(* IEC 61131-3 sources: llm-plc-st-eval/data/definitivo/qwen2.5-coder_14b/I5/zero_shot, 3 files *)

(* ---- ejec_1.st ---- *)
```pascal
FUNCTION_BLOCK FB_Clasificadora
VAR_INPUT
    sensorPresencia : BOOL; // Sensor de presencia de pieza
    sensorAltura : BOOL;    // Sensor de altura de pieza
END_VAR

VAR_OUTPUT
    banda : BOOL;          // Salida para activar la banda
    piston : BOOL;         // Salida para activar el pistón
END_VAR

VAR
    nAltas : INT := 0;      // Contador de piezas altas
    nBajas : INT := 0;      // Contador de piezas bajas
    timer1 : TON;           // Timer para el tiempo de espera (2s)
    timer2 : TON;           // Timer para el tiempo de activación del pistón (1s)
    estado : INT := 0;      // Estado de la máquina de estados
END_VAR

// Máquina de estados
CASE estado OF
    0: // Estado inicial
        banda := TRUE; // La banda funciona continuamente
        IF sensorPresencia THEN
            estado := 1; // Detectada pieza, iniciar temporizador
            timer1(IN := TRUE, PT := T#2S); // Iniciar temporizador de 2s
        END_IF

    1: // Esperando que la pieza llegue al desviador
        IF timer1.Q THEN
            IF sensorAltura THEN
                estado := 2; // Pieza alta, activar pistón
                timer2(IN := TRUE, PT := T#1S); // Iniciar temporizador de 1s
                nAltas := nAltas + 1; // Incrementar contador de piezas altas
            ELSE
                estado := 0; // Pieza baja, continuar
                nBajas := nBajas + 1; // Incrementar contador de piezas bajas
            END_IF
        END_IF

    2: // Activando el pistón
        piston := TRUE;
        IF timer2.Q THEN
            piston := FALSE; // Desactivar pistón
            estado := 0; // Volver al estado inicial
        END_IF

    ELSE
        estado := 0; // Estado desconocido, volver al inicial
END_CASE
```

(* ---- ejec_2.st ---- *)
```iec
FUNCTION_BLOCK FB_Clasificadora
VAR_INPUT
    sensorPresencia : BOOL; // Sensor de presencia de pieza
    sensorAltura : BOOL;    // Sensor de altura de pieza
END_VAR

VAR_OUTPUT
    banda : BOOL;          // Salida para activar la banda
    piston : BOOL;         // Salida para activar el pistón
    nAltas : INT;          // Contador de piezas altas
    nBajas : INT;          // Contador de piezas bajas
END_VAR

VAR
    timer1 : TON;           // Timer para esperar 2 segundos
    timer2 : TON;           // Timer para activar el pistón durante 1 segundo
    piezaDetectada : BOOL;  // Bandera para detectar pieza
END_VAR

// Inicialización de variables
IF NOT piezaDetectada THEN
    timer1(IN := FALSE);
    timer2(IN := FALSE);
    piston := FALSE;
END_IF

// Detectar pieza
IF sensorPresencia AND NOT piezaDetectada THEN
    piezaDetectada := TRUE;
    timer1(IN := TRUE);
    timer1(PTR := T#2S);
END_IF

// Esperar 2 segundos antes de evaluar la altura
IF timer1.Q THEN
    timer1(IN := FALSE);
    IF sensorAltura THEN
        nAltas := nAltas + 1;
        timer2(IN := TRUE);
        timer2(PTR := T#1S);
        piston := TRUE;
    ELSE
        nBajas := nBajas + 1;
    END_IF
END_IF

// Activar el pistón durante 1 segundo
IF timer2.Q THEN
    timer2(IN := FALSE);
    piston := FALSE;
END_IF

// Mantener la banda activa
banda := TRUE;

// Reiniciar la bandera de detección de pieza
IF sensorPresencia = FALSE THEN
    piezaDetectada := FALSE;
END_IF
END_FUNCTION_BLOCK
```

(* ---- ejec_3.st ---- *)
```iec
FUNCTION_BLOCK FB_Clasificadora
VAR_INPUT
    sensorPresencia : BOOL; // Sensor de presencia de pieza
    sensorAltura : BOOL; // Sensor de altura de pieza
END_VAR

VAR_OUTPUT
    banda : BOOL; // Salida de la banda transportadora
    piston : BOOL; // Salida del pistón para desviar piezas altas
    nAltas : INT; // Contador de piezas altas
    nBajas : INT; // Contador de piezas bajas
END_VAR

VAR
    timerDelay : TON; // Temporizador para el retardo de 2 segundos
    timerPiston : TON; // Temporizador para el activo del pistón durante 1 segundo
    piezaDetectada : BOOL; // Bandera para indicar si una pieza ha sido detectada
END_VAR

// Inicialización de temporizadores
timerDelay(IN := FALSE, PT := T#2S);
timerPiston(IN := FALSE, PT := T#1S);

// Banda transportadora siempre activa
banda := TRUE;

// Proceso principal
IF sensorPresencia THEN
    piezaDetectada := TRUE;
    timerDelay(IN := TRUE); // Iniciar el temporizador de retardo
ELSEIF piezaDetectada THEN
    IF timerDelay.Q THEN
        IF sensorAltura THEN
            nAltas := nAltas + 1; // Incrementar contador de piezas altas
            timerPiston(IN := TRUE); // Iniciar el temporizador del pistón
            piston := TRUE; // Activar el pistón
        ELSE
            nBajas := nBajas + 1; // Incrementar contador de piezas bajas
        END_IF
        piezaDetectada := FALSE; // Resetear la bandera de detección
    END_IF
END_IF

// Control del pistón
IF timerPiston.Q THEN
    timerPiston(IN := FALSE); // Detener el temporizador del pistón
    piston := FALSE; // Desactivar el pistón
END_IF
END_FUNCTION_BLOCK
```
